// TIA Portal V17 export
FUNCTION "MCP_RC_FC" : Void   // FC, SCL
BEGIN
END_FUNCTION
